(* Logix 5000 project; controller TFF vendor 1 type 14 code 107 rev 34.11; software revision 34.03; part 36 of 36 *)
(* tags used below, declared in another part *)
   Index : DINT;   // Index
   Index2 : DINT;   // Index
   Index3 : DINT;   // Index
   FlowPath : FlowPath[64];   // Flow Path Array
   FlowPathControl : FlowPathControl;   // Flow Path Control
   FlowPathSetup : FlowPathSetup;   // Flow Path Setup Data
   Valve : Valve[100];   // Valve Array
   ValveControl : ValveControl;   // Valve Control
(* Process, continued *)

ROUTINE Valve_FlowPath   (* ladder *)
// Flow Path Routine
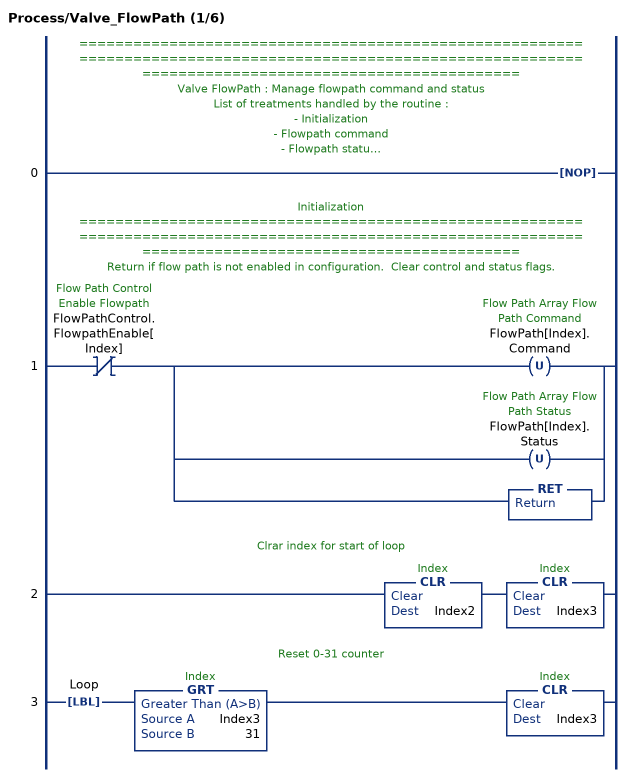
   // ==========================================================================================================================================================
   //                                                                                                  Valve FlowPath : Manage flowpath command and status
   //                                                     List of treatments handled by the routine :
   //                                                          - Initialization
   //                                                          - Flowpath command
   //                                                          - Flowpath status
   //                                                          - Reset flowpath command
   //                                                     -----------------------------------------------------------------------------------------------------------------------------------------------------
   //                                                     History
   //                                                          2019-AUG-13 - Actemium - B. Roch - Initial version for Candidate Release 3.00.00.00.a
   // ========================================================================================================================================================
   0: NOP();
   // Initialization
   // ==========================================================================================================================================================
   // Return if flow path is not enabled in configuration.  Clear control and status flags.
   1: XIO(FlowPathControl.FlowpathEnable[Index])[OTU(FlowPath[Index].Command) ,OTU(FlowPath[Index].Status) ,RET() ];
   // Clrar index for start of loop
   2: CLR(Index2)CLR(Index3);
   // Reset 0-31 counter
   3: LBL(Loop)GRT(Index3,31)CLR(Index3);
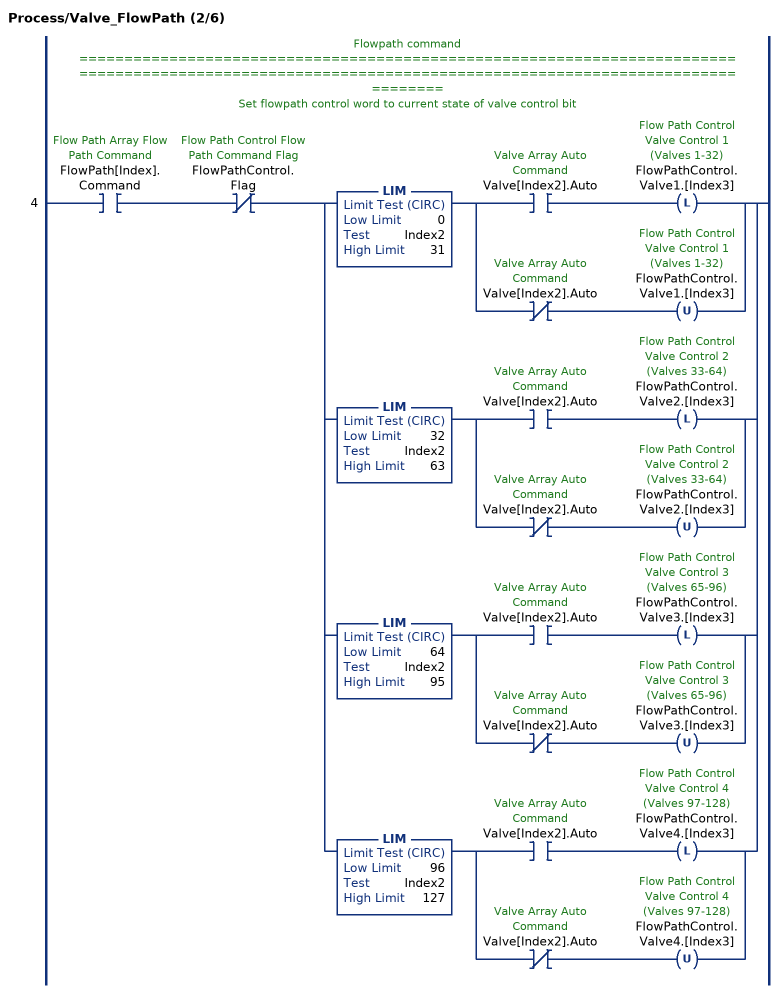
   // Flowpath command
   // ==========================================================================================================================================================
   // Set flowpath control word to current state of valve control bit
   4: XIC(FlowPath[Index].Command)XIO(FlowPathControl.Flag)[LIM(0,Index2,31) [XIC(Valve[Index2].Auto) OTL(FlowPathControl.Valve1.[Index3]) ,XIO(Valve[Index2].Auto) OTU(FlowPathControl.Valve1.[Index3]) ] ,LIM(32,Index2,63) [XIC(Valve[Index2].Auto) OTL(FlowPathControl.Valve2.[Index3]) ,XIO(Valve[Index2].Auto) OTU(FlowPathControl.Valve2.[Index3]) ] ,LIM(64,Index2,95) [XIC(Valve[Index2].Auto) OTL(FlowPathControl.Valve3.[Index3]) ,XIO(Valve[Index2].Auto) OTU(FlowPathControl.Valve3.[Index3]) ] ,LIM(96,Index2,127) [XIC(Valve[Index2].Auto) OTL(FlowPathControl.Valve4.[Index3]) ,XIO(Valve[Index2].Auto) OTU(FlowPathControl.Valve4.[Index3]) ] ];
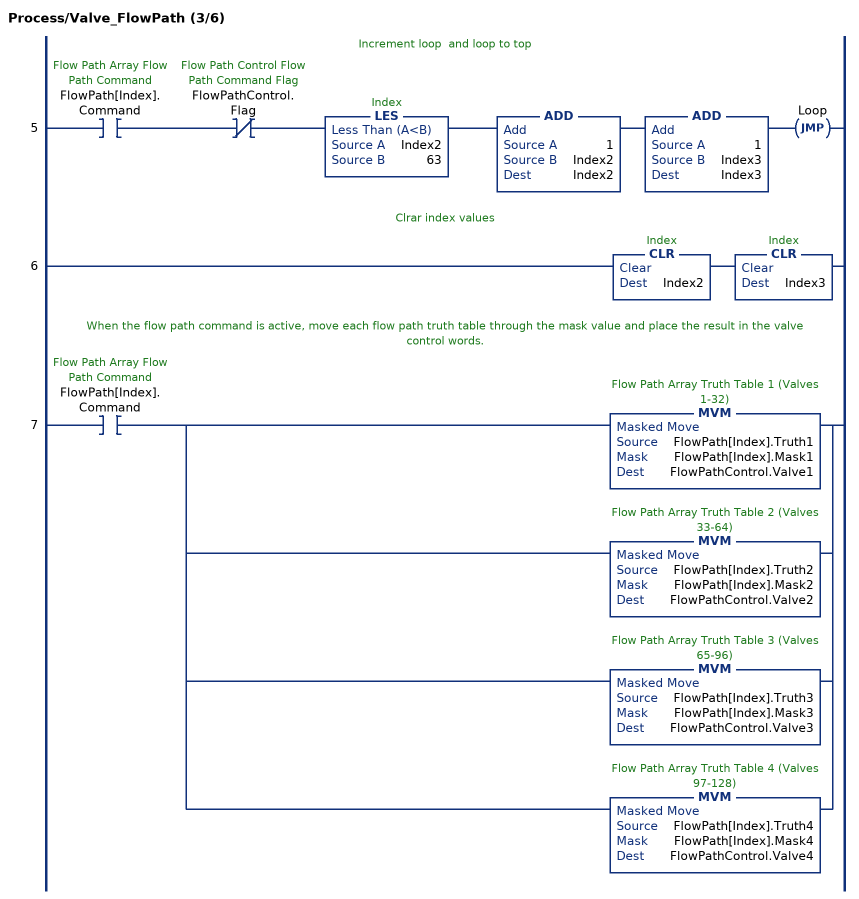
   // Increment loop  and loop to top
   5: XIC(FlowPath[Index].Command)XIO(FlowPathControl.Flag)LES(Index2,63)ADD(1,Index2,Index2)ADD(1,Index3,Index3)JMP(Loop);
   // Clrar index values
   6: CLR(Index2)CLR(Index3);
   // When the flow path command is active, move each flow path truth table through the mask value and place the result in the valve control words.
   7: XIC(FlowPath[Index].Command)[MVM(FlowPath[Index].Truth1,FlowPath[Index].Mask1,FlowPathControl.Valve1) ,MVM(FlowPath[Index].Truth2,FlowPath[Index].Mask2,FlowPathControl.Valve2) ,MVM(FlowPath[Index].Truth3,FlowPath[Index].Mask3,FlowPathControl.Valve3) ,MVM(FlowPath[Index].Truth4,FlowPath[Index].Mask4,FlowPathControl.Valve4) ];
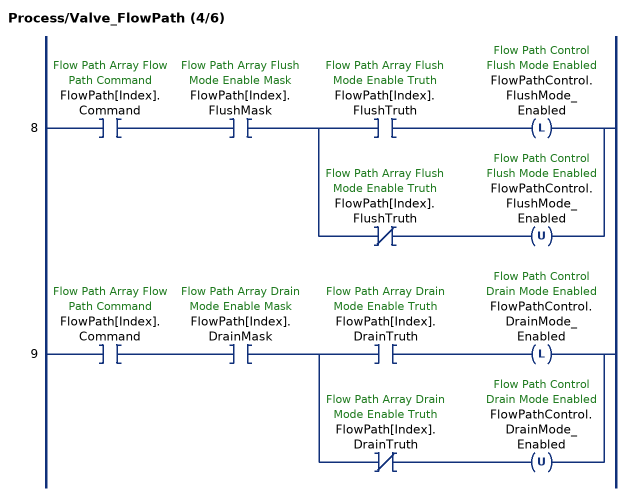
   8: XIC(FlowPath[Index].Command)XIC(FlowPath[Index].FlushMask)[XIC(FlowPath[Index].FlushTruth) OTL(FlowPathControl.FlushMode_Enabled) ,XIO(FlowPath[Index].FlushTruth) OTU(FlowPathControl.FlushMode_Enabled) ];
   9: XIC(FlowPath[Index].Command)XIC(FlowPath[Index].DrainMask)[XIC(FlowPath[Index].DrainTruth) OTL(FlowPathControl.DrainMode_Enabled) ,XIO(FlowPath[Index].DrainTruth) OTU(FlowPathControl.DrainMode_Enabled) ];
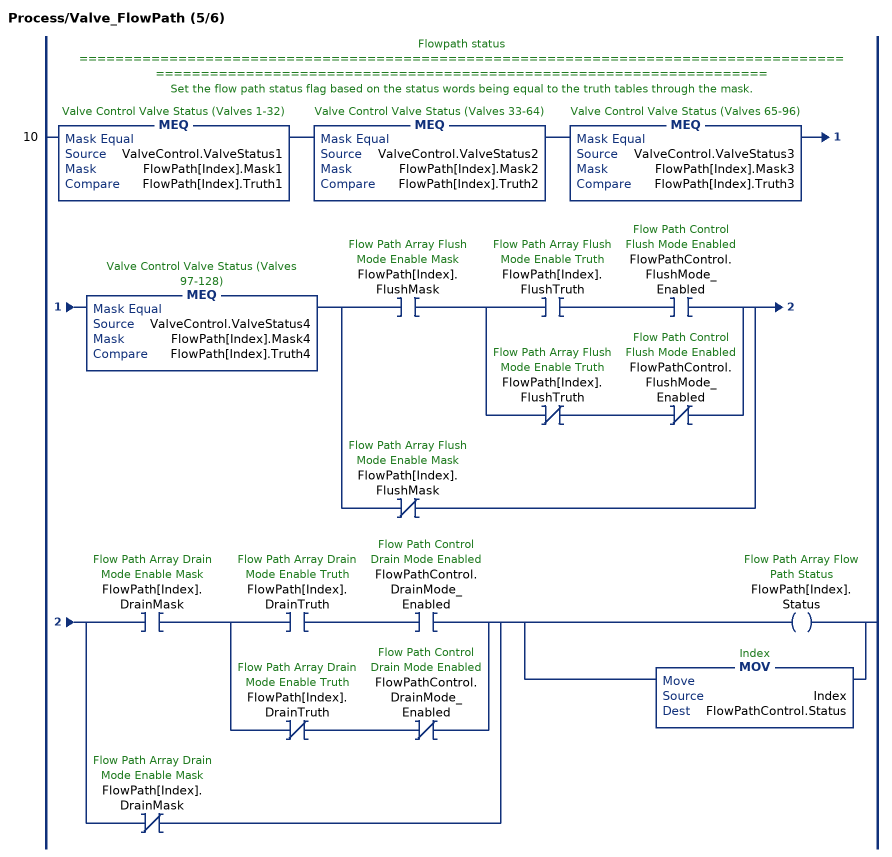
   // Flowpath status
   // =========================================================================================================================================================
   // Set the flow path status flag based on the status words being equal to the truth tables through the mask.
   10: MEQ(ValveControl.ValveStatus1,FlowPath[Index].Mask1,FlowPath[Index].Truth1)MEQ(ValveControl.ValveStatus2,FlowPath[Index].Mask2,FlowPath[Index].Truth2)MEQ(ValveControl.ValveStatus3,FlowPath[Index].Mask3,FlowPath[Index].Truth3)MEQ(ValveControl.ValveStatus4,FlowPath[Index].Mask4,FlowPath[Index].Truth4)[XIC(FlowPath[Index].FlushMask) [XIC(FlowPath[Index].FlushTruth) XIC(FlowPathControl.FlushMode_Enabled) ,XIO(FlowPath[Index].FlushTruth) XIO(FlowPathControl.FlushMode_Enabled) ] ,XIO(FlowPath[Index].FlushMask) ][XIC(FlowPath[Index].DrainMask) [XIC(FlowPath[Index].DrainTruth) XIC(FlowPathControl.DrainMode_Enabled) ,XIO(FlowPath[Index].DrainTruth) XIO(FlowPathControl.DrainMode_Enabled) ] ,XIO(FlowPath[Index].DrainMask) ][OTE(FlowPath[Index].Status) ,MOV(Index,FlowPathControl.Status) ];
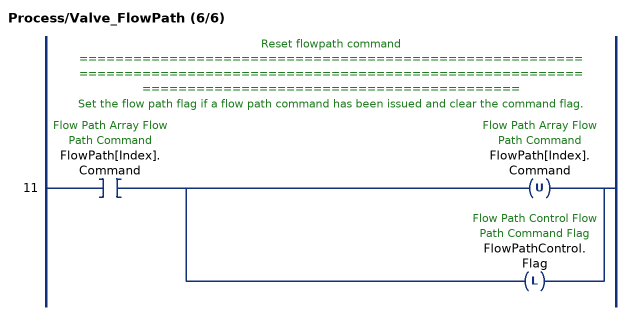
   // Reset flowpath command
   // ==========================================================================================================================================================
   // Set the flow path flag if a flow path command has been issued and clear the command flag.
   11: XIC(FlowPath[Index].Command)[OTU(FlowPath[Index].Command) ,OTL(FlowPathControl.Flag) ];
END_ROUTINE

ROUTINE Valve_FlowPathSetup   (* ladder *)
// Flow Path Setup Routine
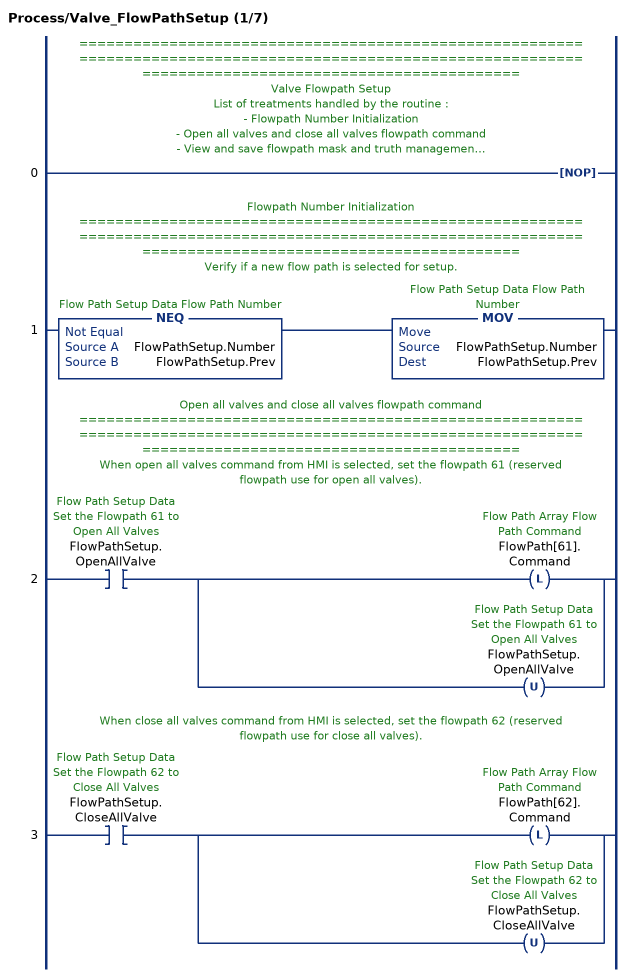
   // ==========================================================================================================================================================
   //                                                                                                                           Valve Flowpath Setup
   //                                                     List of treatments handled by the routine :
   //                                                          - Flowpath Number Initialization
   //                                                          - Open all valves and close all valves flowpath command
   //                                                          - View and save flowpath mask and truth management
   //                                                          - Apply, view mask and view truth command management
   //                                                     -----------------------------------------------------------------------------------------------------------------------------------------------------
   //                                                     History
   //                                                          2019-AUG-13 - Actemium - B. Roch - Initial version for Candidate Release 3.00.00.00.a
   // ==========================================================================================================================================================
   0: NOP();
   // Flowpath Number Initialization
   // ==========================================================================================================================================================
   // Verify if a new flow path is selected for setup.
   1: NEQ(FlowPathSetup.Number,FlowPathSetup.Prev)MOV(FlowPathSetup.Number,FlowPathSetup.Prev);
   // Open all valves and close all valves flowpath command
   // ==========================================================================================================================================================
   // When open all valves command from HMI is selected, set the flowpath 61 (reserved flowpath use for open all valves).
   2: XIC(FlowPathSetup.OpenAllValve)[OTL(FlowPath[61].Command) ,OTU(FlowPathSetup.OpenAllValve) ];
   // When close all valves command from HMI is selected, set the flowpath 62 (reserved flowpath use for close all valves).
   3: XIC(FlowPathSetup.CloseAllValve)[OTL(FlowPath[62].Command) ,OTU(FlowPathSetup.CloseAllValve) ];
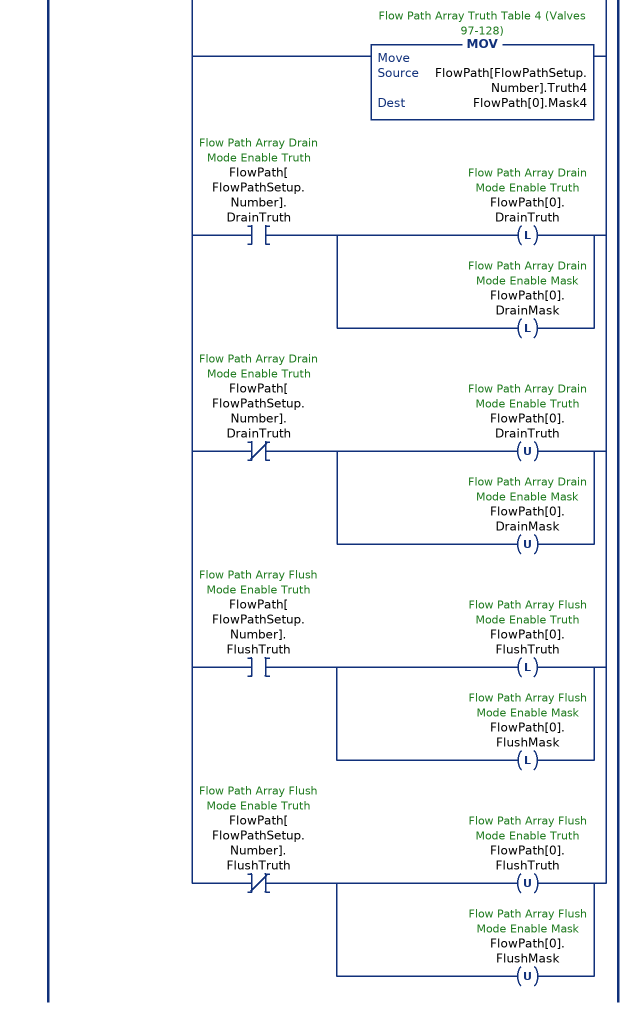
   // View and save flowpath mask and truth management
   // ==========================================================================================================================================================
   // When view truth command from the HMI is set, copy the truth tables of selected flowpath to the truth and mask tables of flowpath 0 (reserved flowpath use for configuration).
   4: XIC(FlowPathSetup.Truth_View)[MOV(FlowPath[FlowPathSetup.Number].Truth1,FlowPath[0].Truth1) ,MOV(FlowPath[FlowPathSetup.Number].Truth1,FlowPath[0].Mask1) ,MOV(FlowPath[FlowPathSetup.Number].Truth2,FlowPath[0].Truth2) ,MOV(FlowPath[FlowPathSetup.Number].Truth2,FlowPath[0].Mask2) ,MOV(FlowPath[FlowPathSetup.Number].Truth3,FlowPath[0].Truth3) ,MOV(FlowPath[FlowPathSetup.Number].Truth3,FlowPath[0].Mask3) ,MOV(FlowPath[FlowPathSetup.Number].Truth4,FlowPath[0].Truth4) ,MOV(FlowPath[FlowPathSetup.Number].Truth4,FlowPath[0].Mask4) ,[XIC(FlowPath[FlowPathSetup.Number].DrainTruth) [OTL(FlowPath[0].DrainTruth) ,OTL(FlowPath[0].DrainMask) ] ,XIO(FlowPath[FlowPathSetup.Number].DrainTruth) [OTU(FlowPath[0].DrainTruth) ,OTU(FlowPath[0].DrainMask) ] ] ,[XIC(FlowPath[FlowPathSetup.Number].FlushTruth) [OTL(FlowPath[0].FlushTruth) ,OTL(FlowPath[0].FlushMask) ] ,XIO(FlowPath[FlowPathSetup.Number].FlushTruth) [OTU(FlowPath[0].FlushTruth) ,OTU(FlowPath[0].FlushMask) ] ] ];
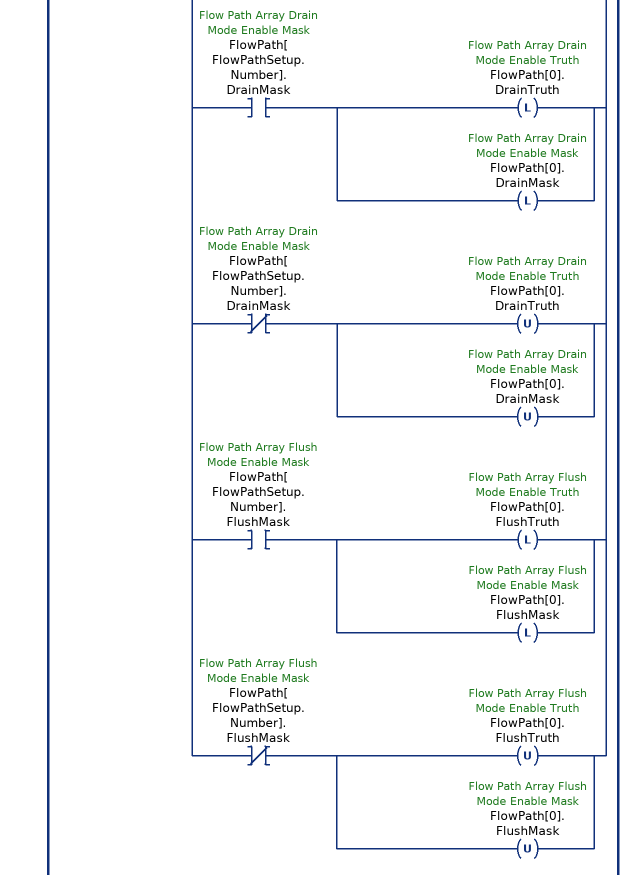
   // When view mask command from the HMI is set, copy the mask tables of selected flowpath to the truth and mask tables of flowpath 0 (reserved flowpath use for configuration).
   5: XIC(FlowPathSetup.Mask_View)[MOV(FlowPath[FlowPathSetup.Number].Mask1,FlowPath[0].Truth1) ,MOV(FlowPath[FlowPathSetup.Number].Mask1,FlowPath[0].Mask1) ,MOV(FlowPath[FlowPathSetup.Number].Mask2,FlowPath[0].Truth2) ,MOV(FlowPath[FlowPathSetup.Number].Mask2,FlowPath[0].Mask2) ,MOV(FlowPath[FlowPathSetup.Number].Mask3,FlowPath[0].Truth3) ,MOV(FlowPath[FlowPathSetup.Number].Mask3,FlowPath[0].Mask3) ,MOV(FlowPath[FlowPathSetup.Number].Mask4,FlowPath[0].Truth4) ,MOV(FlowPath[FlowPathSetup.Number].Mask4,FlowPath[0].Mask4) ,[XIC(FlowPath[FlowPathSetup.Number].DrainMask) [OTL(FlowPath[0].DrainTruth) ,OTL(FlowPath[0].DrainMask) ] ,XIO(FlowPath[FlowPathSetup.Number].DrainMask) [OTU(FlowPath[0].DrainTruth) ,OTU(FlowPath[0].DrainMask) ] ] ,[XIC(FlowPath[FlowPathSetup.Number].FlushMask) [OTL(FlowPath[0].FlushTruth) ,OTL(FlowPath[0].FlushMask) ] ,XIO(FlowPath[FlowPathSetup.Number].FlushMask) [OTU(FlowPath[0].FlushTruth) ,OTU(FlowPath[0].FlushMask) ] ] ];
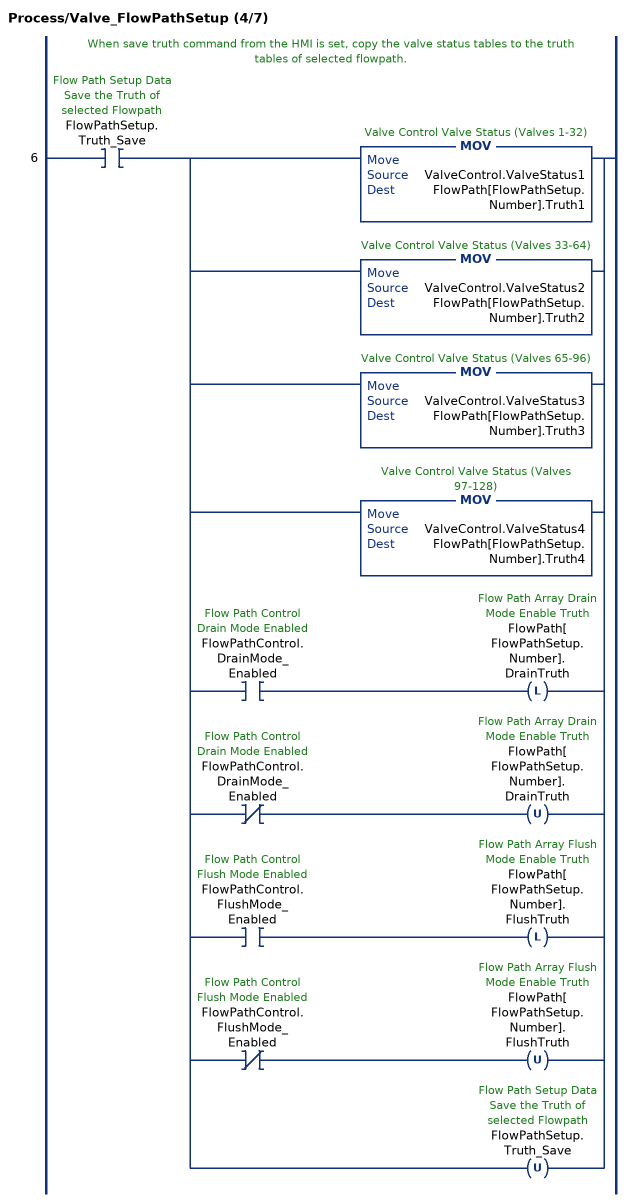
   // When save truth command from the HMI is set, copy the valve status tables to the truth tables of selected flowpath.
   6: XIC(FlowPathSetup.Truth_Save)[MOV(ValveControl.ValveStatus1,FlowPath[FlowPathSetup.Number].Truth1) ,MOV(ValveControl.ValveStatus2,FlowPath[FlowPathSetup.Number].Truth2) ,MOV(ValveControl.ValveStatus3,FlowPath[FlowPathSetup.Number].Truth3) ,MOV(ValveControl.ValveStatus4,FlowPath[FlowPathSetup.Number].Truth4) ,[XIC(FlowPathControl.DrainMode_Enabled) OTL(FlowPath[FlowPathSetup.Number].DrainTruth) ,XIO(FlowPathControl.DrainMode_Enabled) OTU(FlowPath[FlowPathSetup.Number].DrainTruth) ] ,[XIC(FlowPathControl.FlushMode_Enabled) OTL(FlowPath[FlowPathSetup.Number].FlushTruth) ,XIO(FlowPathControl.FlushMode_Enabled) OTU(FlowPath[FlowPathSetup.Number].FlushTruth) ] ,OTU(FlowPathSetup.Truth_Save) ];
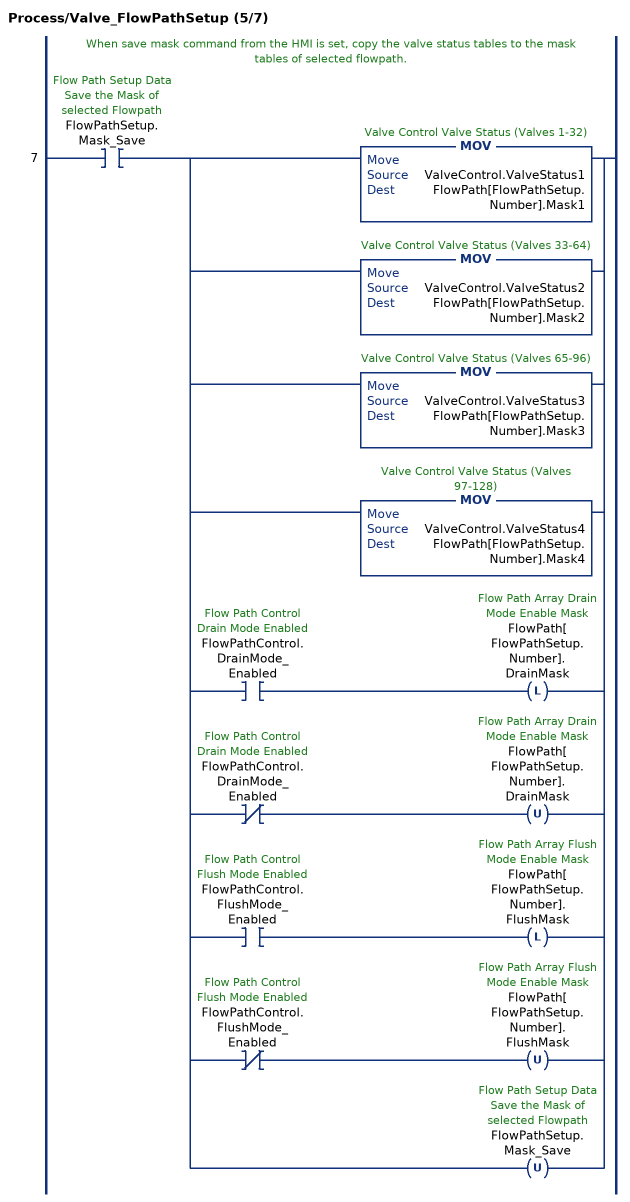
   // When save mask command from the HMI is set, copy the valve status tables to the mask tables of selected flowpath.
   7: XIC(FlowPathSetup.Mask_Save)[MOV(ValveControl.ValveStatus1,FlowPath[FlowPathSetup.Number].Mask1) ,MOV(ValveControl.ValveStatus2,FlowPath[FlowPathSetup.Number].Mask2) ,MOV(ValveControl.ValveStatus3,FlowPath[FlowPathSetup.Number].Mask3) ,MOV(ValveControl.ValveStatus4,FlowPath[FlowPathSetup.Number].Mask4) ,[XIC(FlowPathControl.DrainMode_Enabled) OTL(FlowPath[FlowPathSetup.Number].DrainMask) ,XIO(FlowPathControl.DrainMode_Enabled) OTU(FlowPath[FlowPathSetup.Number].DrainMask) ] ,[XIC(FlowPathControl.FlushMode_Enabled) OTL(FlowPath[FlowPathSetup.Number].FlushMask) ,XIO(FlowPathControl.FlushMode_Enabled) OTU(FlowPath[FlowPathSetup.Number].FlushMask) ] ,OTU(FlowPathSetup.Mask_Save) ];
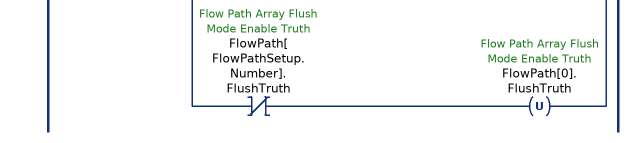
   // Apply, view mask and view truth command management
   // ==========================================================================================================================================================
   // When the flow path applied command from the HMI is set, copy the mask and truth tables of selected flowpath to the flow path 0 mask and truth tables.
   8: XIC(FlowPathSetup.Apply)[MOV(FlowPath[FlowPathSetup.Number].Mask1,FlowPath[0].Mask1) ,MOV(FlowPath[FlowPathSetup.Number].Truth1,FlowPath[0].Truth1) ,MOV(FlowPath[FlowPathSetup.Number].Mask2,FlowPath[0].Mask2) ,MOV(FlowPath[FlowPathSetup.Number].Truth2,FlowPath[0].Truth2) ,MOV(FlowPath[FlowPathSetup.Number].Mask3,FlowPath[0].Mask3) ,MOV(FlowPath[FlowPathSetup.Number].Truth3,FlowPath[0].Truth3) ,MOV(FlowPath[FlowPathSetup.Number].Mask4,FlowPath[0].Mask4) ,MOV(FlowPath[FlowPathSetup.Number].Truth4,FlowPath[0].Truth4) ,[XIC(FlowPath[FlowPathSetup.Number].DrainMask) OTL(FlowPath[0].DrainMask) ,XIO(FlowPath[FlowPathSetup.Number].DrainMask) OTU(FlowPath[0].DrainMask) ] ,[XIC(FlowPath[FlowPathSetup.Number].FlushMask) OTL(FlowPath[0].FlushMask) ,XIO(FlowPath[FlowPathSetup.Number].FlushMask) OTU(FlowPath[0].FlushMask) ] ,[XIC(FlowPath[FlowPathSetup.Number].DrainTruth) OTL(FlowPath[0].DrainTruth) ,XIO(FlowPath[FlowPathSetup.Number].DrainTruth) OTU(FlowPath[0].DrainTruth) ] ,[XIC(FlowPath[FlowPathSetup.Number].FlushTruth) OTL(FlowPath[0].FlushTruth) ,XIO(FlowPath[FlowPathSetup.Number].FlushTruth) OTU(FlowPath[0].FlushTruth) ] ];
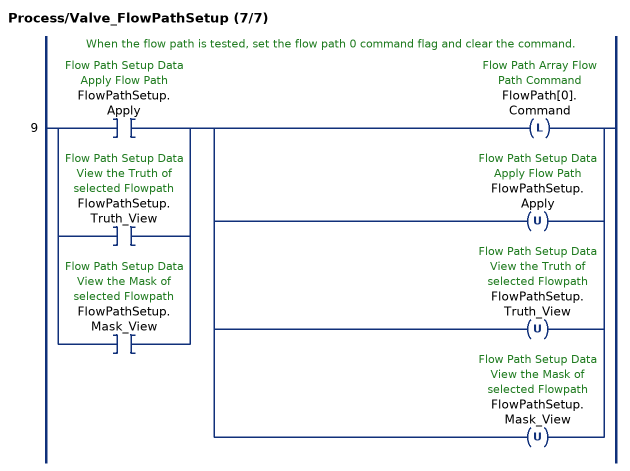
   // When the flow path is tested, set the flow path 0 command flag and clear the command.
   9: [XIC(FlowPathSetup.Apply) ,XIC(FlowPathSetup.Truth_View) ,XIC(FlowPathSetup.Mask_View) ][OTL(FlowPath[0].Command) ,OTU(FlowPathSetup.Apply) ,OTU(FlowPathSetup.Truth_View) ,OTU(FlowPathSetup.Mask_View) ];
END_ROUTINE
END_PROGRAM
